// TIA Portal V19 export
TYPE "ST_TPM_AutoPosition"
   STRUCT
      X : Int;
      Y : Int;
      Z : Int;
      Rx : Int;
      Ry : Int;
      Rz : Int;
   END_STRUCT;
END_TYPE
